(* IEC 61131-3 sources: llm-plc-st-eval/data/processed_definitivo/qwen2.5-coder_14b/A5/few_shot, 3 files *)

(* ---- ejec_1.st ---- *)
FUNCTION_BLOCK FB_Registro
VAR_INPUT
    evento : INT; (* Código del evento *)
    nuevoEvento : BOOL; (* Indica si se ha producido un nuevo evento *)
    ciclo : TIME; (* Tiempo de ciclo de ejecución *)
END_VAR
VAR_OUTPUT
    buffer : ARRAY[0..19] OF ST_Evento; (* Buffer de eventos *)
    indice : INT; (* Índice del último evento registrado *)
    nEventos : INT; (* Número de eventos válidos en el buffer *)
END_VAR
VAR
    tiempoAcumulado : TIME := T#0s; (* Tiempo acumulado desde el arranque *)
    eventoAnterior : BOOL := FALSE; (* Estado anterior de nuevoEvento *)
END_VAR

(* Definición de la estructura ST_Evento *)
TYPE ST_Evento :
    STRUCT
        codigo : INT; (* Código del evento *)
        marca : TIME; (* Marca de tiempo del evento *)
    END_STRUCT
END_TYPE

(* Acumulación del tiempo *)
tiempoAcumulado := tiempoAcumulado + ciclo;

(* Registro de eventos *)
IF nuevoEvento AND NOT eventoAnterior THEN
    IF indice = -1 THEN
        indice := 0;
    ELSE
        indice := (indice + 1) MOD 20;
    END_IF

    buffer[indice].codigo := evento;
    buffer[indice].marca := tiempoAcumulado;

    IF nEventos < 20 THEN
        nEventos := nEventos + 1;
    END_IF
END_IF

(* Actualización del estado anterior de nuevoEvento *)
eventoAnterior := nuevoEvento;
END_FUNCTION_BLOCK

(* ---- ejec_2.st ---- *)
TYPE ST_Evento :
STRUCT
    codigo : INT; (* Código del evento *)
    marca : TIME; (* Marca de tiempo del evento *)
END_STRUCT
END_TYPE

FUNCTION_BLOCK FB_Registro
VAR_INPUT
    evento : INT; (* Código del evento *)
    nuevoEvento : BOOL; (* Indica si se debe registrar un nuevo evento *)
    ciclo : TIME; (* Período de ejecución del bloque *)
END_VAR
VAR_OUTPUT
    buffer : ARRAY[0..19] OF ST_Evento; (* Buffer de eventos *)
    indice : INT; (* Índice del último evento registrado *)
    nEventos : INT; (* Número de eventos válidos en el buffer *)
END_VAR
VAR
    tiempoAcumulado : TIME := T#0s; (* Tiempo acumulado desde el arranque *)
    ultimoEvento : INT := -1; (* Índice del último evento registrado *)
    eventosRegistrados : INT := 0; (* Número de eventos registrados *)
END_VAR

(* Acumula el tiempo de ciclo *)
tiempoAcumulado := tiempoAcumulado + ciclo;

(* Registro de nuevo evento *)
IF nuevoEvento THEN
    (* Incrementa el índice y ajusta si se llena el buffer *)
    ultimoEvento := (ultimoEvento + 1) MOD 20;

    (* Registra el evento en el buffer *)
    buffer[ultimoEvento].codigo := evento;
    buffer[ultimoEvento].marca := tiempoAcumulado;

    (* Actualiza el número de eventos válidos *)
    IF eventosRegistrados < 20 THEN
        eventosRegistrados := eventosRegistrados + 1;
    END_IF;

    (* Actualiza el índice y el número de eventos *)
    indice := ultimoEvento;
    nEventos := eventosRegistrados;
END_IF
END_FUNCTION_BLOCK

(* ---- ejec_3.st ---- *)
FUNCTION_BLOCK FB_Registro
VAR_INPUT
    evento : INT; (* Código del evento *)
    nuevoEvento : BOOL; (* Indica si se debe registrar un nuevo evento *)
    ciclo : TIME; (* Período de ejecución del bloque *)
END_VAR
VAR_OUTPUT
    buffer : ARRAY[0..19] OF ST_Evento; (* Buffer circular de eventos *)
    indice : INT; (* Índice de la posición del último evento registrado *)
    nEventos : INT; (* Número de eventos válidos en el buffer *)
END_VAR
VAR
    tiempoAcumulado : TIME := T#0s; (* Tiempo acumulado desde el arranque *)
    eventoAnterior : BOOL := FALSE; (* Estado anterior de nuevoEvento *)
END_VAR

(* Definición de la estructura ST_Evento *)
TYPE ST_Evento :
STRUCT
    codigo : INT; (* Código del evento *)
    marca : TIME; (* Marca de tiempo del evento *)
END_STRUCT
END_TYPE

(* Acumulación del tiempo *)
tiempoAcumulado := tiempoAcumulado + ciclo;

(* Registro de nuevo evento *)
IF nuevoEvento AND NOT eventoAnterior THEN
    (* Incrementar el índice y ajustarlo al rango del buffer *)
    indice := (indice + 1) MOD 20;

    (* Registrar el evento en el buffer *)
    buffer[indice].codigo := evento;
    buffer[indice].marca := tiempoAcumulado;

    (* Actualizar el número de eventos válidos *)
    IF nEventos < 20 THEN
        nEventos := nEventos + 1;
    END_IF;
END_IF;

(* Actualizar el estado anterior de nuevoEvento *)
eventoAnterior := nuevoEvento;
END_FUNCTION_BLOCK
